FUNCTION_BLOCK "640_Rollenbahnen"   // FB640, SCL
{ S7_Optimized_Access := 'FALSE' }
AUTHOR : DJonas
VERSION : 0.1
   VAR_INPUT
      Notaus : Bool;
      Betriebsbereit : Bool;
      Start : Bool;
      StartRB : Bool;
      "630_Grundstellung" : Bool;
      i_s_grün : Bool;
      i_s_blau : Bool;
      i_Farbe_Code : Int;
   END_VAR
   VAR_OUTPUT
      o_RB_Frei : Bool;
      o_kontrolliert : Bool;
   END_VAR
   VAR_IN_OUT
      o_Farbsensor_Code : Int;
      o_kontrolle_fehler : Bool;
   END_VAR
   VAR
      RB9001_belegt : Bool;
      RB9002_belegt : Bool;
      RB9003_Belegt : Bool;
      Fehler : Bool;
      Neustart : TP;
      RB9001 : "641_Rollenbahn";
      RB9002 : "641_Rollenbahn";
      RB9003 : "641_Rollenbahn";
      B9002_RB9001_ntrig : "1001_300-ntrig-scl";
      B9004_RB9002_ntrig : "1001_300-ntrig-scl";
      B9006_RB9003_ntrig : "1001_300-ntrig-scl";
   END_VAR
BEGIN
   // Neustart Rollenbahn 2s laufen lassen um evtl. vorhandene Paletten vor einen Sensor zu fördern
   #Neustart(IN := #Notaus AND #Betriebsbereit, PT := T#2s);

   // Fehler Überbabe ohne Palette
   IF #StartRB AND NOT ("B9001_RB9001" OR "B9002_RB9001") THEN
       #Fehler := 1;
   ELSIF "B9006_RB9003" THEN
       #Fehler := 0;
   END_IF; 

   // Farbcode der Sensoren erstellen
   IF #i_s_blau THEN
       #o_Farbsensor_Code := 1;
   ELSIF #i_s_grün THEN
       #o_Farbsensor_Code := 2;
   ELSE
       #o_Farbsensor_Code := 0;
   END_IF;

   // Erkennung falsche Farbe auf Palette
   // ((#i_s_blau OR #i_s_grün) AND NOT (#i_Farbe_Code = #o_Farbsensor_Code))
   IF #Fehler AND #Betriebsbereit THEN
       #o_kontrolle_fehler := 1;
   END_IF;
   (*
   IF #o_kontrolle_fehler AND #Start THEN
       #o_Farbsensor_Code := #i_Farbe_Code;
       #o_kontrolliert := 1;
       #o_kontrolle_fehler := 0;
       #o_RB_Frei := 0;
       #Fehler := 0;
       RETURN;
   END_IF; *)

   // Kontrolle OK
   #o_kontrolliert := ((#i_s_blau OR #i_s_grün) AND (#i_Farbe_Code = #o_Farbsensor_Code)) OR #RB9003_Belegt OR #Fehler;

   // trigger für Stop Rollenbahn
   #B9002_RB9001_ntrig(IN := "B9002_RB9001" OR #Neustart.Q);
   #B9004_RB9002_ntrig(IN := "B9004_RB9002" OR #Neustart.Q);
   #B9006_RB9003_ntrig(IN := "B9006_RB9003" OR #Neustart.Q);

   // Ausgabe Rollenbahn 9001 und 9002 frei
   #o_RB_Frei := NOT #RB9001.belegt OR NOT #RB9002.belegt OR NOT #RB9003.belegt ;

   // Ansteuerung Rollenbahnen
   #RB9001(i_Start1:=(#StartRB OR #Neustart.Q),
           i_Start2:=("B9001_RB9001" OR "B9002_RB9001") AND #"630_Grundstellung",
           i_Stop:=#B9002_RB9001_ntrig.OUT OR (NOT #Betriebsbereit AND #"630_Grundstellung"),
           i_Halt:= NOT #"630_Grundstellung",
           i_NotHalt:=#Notaus,
           Output=>"RB9001",
           belegt:=#RB9001_belegt);

   #RB9002(i_Start1 := #Neustart.Q,
           i_Start2 := (("B9002_RB9001" AND #RB9001.Output) OR "B9003_RB9002"),
           i_Stop := #B9004_RB9002_ntrig.OUT OR (NOT #Betriebsbereit AND #"630_Grundstellung" AND #o_RB_Frei),
           i_NotHalt := #Notaus,
           Output => "RB9002",
           belegt := #RB9002_belegt);

   #RB9003(i_Start1:=#Neustart.Q,
           i_Start2:=("B9004_RB9002" OR "B9005_RB9003"),
           i_Stop:=#B9006_RB9003_ntrig.OUT OR (NOT #Betriebsbereit AND #"630_Grundstellung" AND #o_RB_Frei),
           i_NotHalt:=#Notaus,
           Output=>"RB9003",
           belegt:=#RB9003_Belegt);
END_FUNCTION_BLOCK

FUNCTION_BLOCK "641_Rollenbahn"   // FB641, SCL
{ S7_Optimized_Access := 'FALSE' }
VERSION : 0.1
   VAR_INPUT
      i_Start1 : Bool;
      i_Start2 : Bool;
      i_Halt : Bool;
      i_Stop : Bool;
      i_NotHalt : Bool;
   END_VAR
   VAR_OUTPUT
      Output : Bool;
   END_VAR
   VAR_IN_OUT
      belegt : Bool;
   END_VAR
BEGIN

   // Rollenbahn belegt setzen
   IF #i_Start1 OR #i_Start2 THEN
       #belegt := 1;
   END_IF;

   // Rollenbahn belegt entfernen
   IF #i_Stop OR NOT #i_NotHalt THEN
       #belegt := 0;
   END_IF;

   // Ausgang setzen wenn Rollenbahn belegt, kein Halt und kein Nothalt(zusätzlicher Schutz)
   #Output := #belegt AND #i_NotHalt AND  NOT #i_Halt;
END_FUNCTION_BLOCK

FUNCTION_BLOCK "1001_300-ntrig-scl"   // FB1001, SCL
{ S7_Optimized_Access := 'FALSE' }
VERSION : 0.1
   VAR_INPUT
      IN : Bool;
   END_VAR
   VAR_OUTPUT
      OUT : Bool;
   END_VAR
   VAR
      Merker : Bool;
   END_VAR
BEGIN
   #OUT := #Merker AND NOT #IN;
   #Merker := #IN;
END_FUNCTION_BLOCK

// ===== library: MasterCopy "RB_TB_einfach" =====

FUNCTION_BLOCK "RB_TB_einfach"   // FB101, GRAPH
{ S7_Optimized_Access := 'FALSE' }
VERSION : 0.1
// Einfacher Steuerbaustein RB / TB 
// Sensor Anfang / Ende  NO
   VAR_INPUT
      INIT_SQ : Bool := false;   // Kette in Initialzustand versetzen
      A_EIN : Bool;
      A_NOT_HALT : Bool;
      Nachfolgendes_Agg_frei : Bool;
      Sensor_vorheriges_Agg : Bool;
      Sensor_Anfang : Bool;   // Öffner
      Sensor_Ende : Bool;   // Öffner
   END_VAR
   VAR_OUTPUT
      Schritt_Nummer : Int;
      Aggregat : Bool;
      Aggregat_frei : Bool;
   END_VAR
   VAR
      HM_FLAM : Array[1..8] of Bool;
      Flanke : Array[1..8] of Bool;
      HM_Agg_Frei : Bool;
      HM_belegt : Bool;
      SWITCH : Array[0..0] of DWord;
      SW_SQTS : Array[0..6] of Byte;
      SW_ADDR : Word := 16#C;
      G7T_0 : GraphTransition;
      G7S_0 : GraphStep;
      PRE_CRIT : Array[0..1] of DWord;
      POST_CRIT : Array[0..0] of DWord;
      TVX : Array[0..2] of Byte;
      TTX : Array[0..2] of Byte;
      TSX : Array[0..2] of Byte;
      S00X : Array[0..2] of Byte;
      SOFFX : Array[0..2] of Byte;
      SONX : Array[0..2] of Byte;
      SAX : Array[0..2] of Byte;
      SERRX : Array[0..7] of Byte;
      SMX : Array[0..7] of Byte;
      S0X : Array[0..7] of Byte;
      S1X : Array[0..7] of Byte;
      S_DISPLAY : Int;   // Interne Anzeige des Ausgangsparameters S_NO
      S_SEL_OLD : Int;   // Vorheriger Wert an S_SEL
      S_DISPIDX : Byte;   // Index des Schritts, der an S_NO anliegt
      T_DISPIDX : Byte;   // Index der Transition, die an T_NO anliegt
      MOPEDGE : Struct
         AUTO : Bool := false;
         MAN : Bool := false;
         TAP : Bool := false;
         TOP : Bool := false;
         ACK_S : Bool := false;
         REG_S : Bool := false;
         T_PREV : Bool := false;
         T_NEXT : Bool := false;
         LOCK : Bool := false;
         SUP : Bool := false;
         ACKREQ : Bool := false;
         SSKIP : Bool := false;
         OFF : Bool := false;
         INIT : Bool := false;
         HALT : Bool := false;
         TMS_HALT : Bool := false;
         OPS_ZERO : Bool := false;
         SACT_DISP : Bool := false;
         SEF_DISP : Bool := false;
         SALL_DISP : Bool := false;
         S_PREV : Bool := false;
         S_NEXT : Bool := false;
         S_SELOK : Bool := false;
         S_ON : Bool := false;
         S_OFF : Bool := false;
         T_PUSH : Bool := false;
         REG : Bool := false;
         ACK : Bool := false;
         IL_PERM : Bool := false;
         T_PERM : Bool := false;
         ILP_MAN : Bool := false;
      END_STRUCT;
      MOP : Struct   // Betriebsart
         AUTO : Bool := true;   // Zustand: Automatischer Betrieb
         MAN : Bool := false;   // Zustand: Handbetrieb
         TAP : Bool := false;   // Zustand: Halbautomatisch/Weiterschalten mit Transition
         TOP : Bool := false;   // Zustand: Halbautomatisch/Ignoriere Transition
         ACK_S : Bool := false;   // Anforderung: Schritt quittieren, der an Parameter S_NO anliegt
         REG_S : Bool := false;   // Anforderung: Schritt registrieren, der an Parameter S_NO anliegt
         T_PREV : Bool := false;   // Anforderung: Vorherige gültige Transition am Parameter T_NO ausgeben
         T_NEXT : Bool := false;   // Anforderung: Nächste gültige Transition am Parameter T_NO ausgeben
         LOCK : Bool := true;   // Zustand: Interlockbearbeitung aktiviert
         SUP : Bool := true;   // Zustand: Supervisionsbearbeitung aktiviert
         ACKREQ : Bool := false;   // Zustand: Quittierung erforderlich
         SSKIP : Bool := false;   // Zustand: "Schritte überspringen" aktiviert
         OFF : Bool := false;   // Anforderung: Alle Schritte deaktivieren
         INIT : Bool := true;   // Anforderung: Kette in Initialzustand schalten
         HALT : Bool := false;   // Zustand: Kette schaltet nicht weiter
         TMS_HALT : Bool := false;   // Zustand: Alle internen Zeiten angehalten
         OPS_ZERO : Bool := false;   // Zustand: Alle mit N, L, D bearbeitete Operanden auf 0 gesetzt
         SACT_DISP : Bool := true;   // Zustand: Nur aktive Schritte anzeigen
         SEF_DISP : Bool := false;   // Zustand: Nur fehlerhafte und gestörte Schritte anzeigen
         SALL_DISP : Bool := false;   // Zustand: Alle Schritte anzeigen
         S_PREV : Bool := false;   // Anforderung: Vorherigen Schritt am Parameter S_NO ausgeben
         S_NEXT : Bool := false;   // Anforderung: Nächsten Schritt am Parameter S_NO ausgeben
         S_SELOK : Bool := false;   // Anforderung: Schrittnummer, die am Parameter S_SEL anliegt, am Parameter S_NO ausgeben
         S_ON : Bool := false;   // Anforderung: Schritt aktivieren, der am Parameter S_NO anliegt
         S_OFF : Bool := false;   // Anforderung: Schritt deaktivieren, der am Parameter S_NO anliegt
         T_PUSH : Bool := false;   // Anforderung: Schaltfreigabe für Transition
         REG : Bool := false;   // Anforderung: Alle Interlock- und Supervisionsfehler registrieren
         ACK : Bool := false;   // Anforderung: Alle Interlock- und Supervisionsfehler quittieren
         IL_PERM : Bool := false;   // Zustand: Permanente Bearbeitung aller Interlocks
         T_PERM : Bool := false;   // Zustand: Permanente Bearbeitung aller Transitionen
         ILP_MAN : Bool := false;   // Zustand: Permanente Bearbeitung aller Interlocks im Handbetrieb
      END_STRUCT;
      TICKS : Struct   // Zeittakte
         DELTA : Time := T#0ms;   // Zeitdifferenz zwischen zwei Zyklen
         OLD : Time := T#0ms;   // 10 ms Taktzählerstand im letzten Zyklus
         NEW : Time := T#0ms;   // 10 ms Taktzählerstand in diesem Zyklus
      END_STRUCT;
      SQ_FLAGS : Struct   // Kettenmerker
         ERR_FLT : Bool := false;   // Sammelfehler Interlock und Supervision
         ERROR : Bool := false;   // Sammelfehler Interlock
         FAULT : Bool := false;   // Sammelfehler Supervision
         RT_FAIL : Bool := false;   // Laufzeitfehler
         NO_SNO : Bool := false;   // Angeforderte Schrittnummer nicht gefunden
         NF_OFL : Bool := false;   // Überlauf: Zu viele Anforderungen ON oder OFF
         SA_OFL : Bool := false;   // Überlauf: Zu viele Schritte aktiv
         TV_OFL : Bool := false;   // Überlauf: Zu viele gültige Transitionen
         MSG_OFL : Bool := false;   // Überlauf: Nicht genügend Systemressourcen fü ALARM_S
         NO_SWI : Bool := false;   // Nicht Schalten in diesem Zyklus
         CYC_OP : Bool := false;   // Zyklische Bearbeitung der Kette nach Initialisierung
         AS_MSG : Bool := true;   // Meldungen zur Laufzeit durch Anweisung aktiviert oder deaktiviert
         AS_SEND : Bool := false;   // Meldungen von WR_USMSG senden oder nur in Diagnosepuffer eintragen
         SQ_BUSY : Bool := false;   // Interner Flankenmerker für Vorgangsbearbeitung
         SA_BUSY : Bool := false;   // Interner Flankenmerker für Vorgangsbearbeitung
         AS_SIG : Bool := false;   // Flankenmerker für Meldungen von Alarm_S und Alarm_SQ
      END_STRUCT;
      S_PTR : DWord := 16#450;
      S_PTR2 : DWord := 16#0;
      S_PTR3 : DWord := 16#D50;
      S_PTR4 : DWord := 16#D10;
      T_PTR : DWord := 16#CD0;
      C_AR2 : DWord := 16#0;
      M_FBDB : DWord := 16#640000;
      M_SNO : Word := 16#4;
      M_EVID : Word := 16#0;
      M_EVIL : C_Alarm_s;
      M_EVSV : C_Alarm_s;
      M_EV : DWord := 16#C30;
      CRIT : Array[0..31] of Bool;
      S_START : Byte := 16#0;
      S_IDX : Byte := 16#0;
      S_INT : Int := 72;
      S_TMP : Byte := 16#0;
      T_START : Byte := 16#0;
      T_IDX : Byte := 16#0;
      T_TMP : Byte := 16#0;
      T_TMP2 : Byte := 16#00;
      TV_POT : Byte := 16#02;
      RETURN1 : Byte := 16#0;
      RETURN2 : Byte := 16#0;
      SINI : Array[0..2] of Byte;
      LSTT : Array[0..6] of Byte;
      ATAJ : Array[0..6] of Byte;
      ATAB : Array[0..6] of Byte;
      PSTT : Array[0..6] of Byte;
      NSTT : Array[0..6] of Byte;
      ASSJ : Array[0..6] of Byte;
      ASSB : Array[0..6] of Byte;
      PTTS : Array[0..6] of Byte;
      NTTS : Array[0..6] of Byte;
      PRE_CNT : Word := 16#2;
      POST_CNT : Word := 16#1;
      ADR_COND : Word := 16#0;
      MAX_TVAL : Byte := 16#1;
      MAX_SACT : Byte := 16#1;
      MAX_CRIT : Byte := 16#4;
      T_CNT : Byte := 16#6;
      SUP_CNT : Byte := 16#0;
      LOCK_CNT : Byte := 16#5;
      S_CNT : Byte := 16#6;
      SQ_CNT : Byte := 16#1;
      PRS_INPAR : DWord := 16#40000000;
      PRS_OUTPAR : DWord := 16#0;
      GC_FLAGS : Struct
         T_MACH : Byte := 16#EB;
         COND_ED : Byte := 16#E2;
         W_LEVEL : Byte := 16#D5;
         FB_IF : Byte := 16#FA;
         AS_MSG : Word := 16#404;
         SSB : Word := 16#108;
         DILG : Word := 16#27E;
         ADDR_T0 : Word := 16#1A;
         CRIT_AVAIL : Bool := false;
         SSKIP_AVAIL : Bool := true;
         SSKIP_ON : Bool := false;
         ACK_REQ : Bool := false;
         SYNC_AVAIL : Bool := true;
         ILP_MAN : Bool := false;
         SWM_LOCKED : Bool := false;
         SAVE_SW : Bool := true;
      END_STRUCT;
      G7_FBMARK : Byte := 16#3C;
      G7_RELEASE : Byte := 16#3C;
      G7_ID2 : Byte := 16#37;
      G7_ID1 : Byte := 16#47;
   END_VAR
   // SW_SQTS[0] := 16#1;
   // TVX[0] := 16#1;
   // TTX[0] := 16#1;
   // TSX[0] := 16#1;
   // S00X[0] := 16#1;
   // SOFFX[0] := 16#1;
   // SONX[0] := 16#1;
   // SAX[0] := 16#1;
   // SERRX[0] := 16#1;
   // SMX[0] := 16#1;
   // S0X[0] := 16#1;
   // S1X[0] := 16#1;
   // SINI[0] := 16#2;
   // SINI[1] := 16#1;
   // SINI[2] := 0;
   // LSTT[0] := 0;
   // LSTT[1] := 0;
   // LSTT[2] := 0;
   // LSTT[3] := 0;
   // LSTT[4] := 0;
   // LSTT[5] := 0;
   // ATAJ[0] := 0;
   // ATAJ[1] := 16#1;
   // ATAJ[2] := 16#2;
   // ATAJ[3] := 16#3;
   // ATAJ[4] := 16#4;
   // ATAJ[5] := 16#5;
   // ATAB[0] := 0;
   // ATAB[1] := 16#1;
   // ATAB[2] := 16#2;
   // ATAB[3] := 16#3;
   // ATAB[4] := 16#4;
   // ATAB[5] := 16#5;
   // PSTT[0] := 0;
   // PSTT[1] := 16#1;
   // PSTT[2] := 16#2;
   // PSTT[3] := 16#3;
   // PSTT[4] := 16#4;
   // PSTT[5] := 16#5;
   // NSTT[0] := 16#1;
   // NSTT[1] := 16#2;
   // NSTT[2] := 16#3;
   // NSTT[3] := 16#4;
   // NSTT[4] := 16#5;
   // NSTT[5] := 16#6;
   // ASSJ[0] := 0;
   // ASSJ[1] := 16#1;
   // ASSJ[2] := 16#2;
   // ASSJ[3] := 16#3;
   // ASSJ[4] := 16#4;
   // ASSJ[5] := 16#5;
   // ASSB[0] := 0;
   // ASSB[1] := 16#1;
   // ASSB[2] := 16#2;
   // ASSB[3] := 16#3;
   // ASSB[4] := 16#4;
   // ASSB[5] := 16#5;
   // PTTS[0] := 0;
   // PTTS[2] := 16#1;
   // PTTS[3] := 16#2;
   // PTTS[4] := 16#3;
   // PTTS[5] := 16#4;
   // NTTS[0] := 0;
   // NTTS[1] := 16#1;
   // NTTS[2] := 16#2;
   // NTTS[3] := 16#3;
   // NTTS[4] := 16#4;
   // NTTS[5] := 16#5;
   // LSTT[6] := 16#1;
   // ATAJ[6] := 16#6;
   // ATAB[6] := 16#6;
   // PSTT[6] := 16#6;
   // NSTT[6] := 16#1;
   // ASSJ[6] := 16#6;
   // ASSB[6] := 16#6;
   // PTTS[6] := 16#5;
   // NTTS[6] := 16#6;
BEGIN
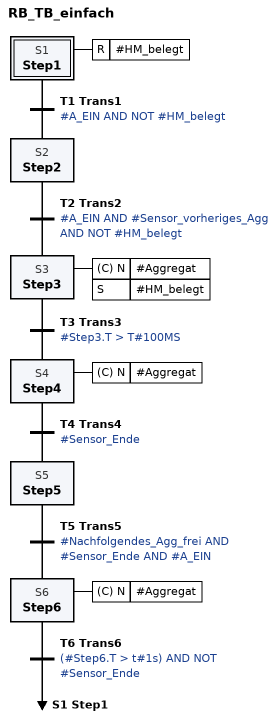
   // permanent pre-instructions
   NETWORK 1
      #HM_Agg_Frei := NOT #HM_belegt;
      #Aggregat_frei := NOT #HM_belegt;
   NETWORK 2
   TITLE = Ausgabe Schrittnummer
      #Schritt_Nummer := #S_DISPLAY;

   // sequencer 1
   INITIAL_STEP Step1:   // S1
      interlock C := NOT #A_NOT_HALT;
      // Warten auf Start
              R    #HM_belegt
   END_STEP
   TRANSITION Trans1 FROM Step1 TO Step2   // T1
      := #A_EIN AND NOT #HM_belegt;
   END_TRANSITION
   STEP Step4:   // S4
      interlock C := NOT #A_NOT_HALT;
      // Einfahrt bis Ende
      (C)     N    #Aggregat
   END_STEP
   TRANSITION Trans4 FROM Step4 TO Step5   // T4
      := #Sensor_Ende;
   END_TRANSITION
   STEP Step5:   // S5
      interlock C := NOT #A_NOT_HALT;
      // Warten auf Ausfahrt
   END_STEP
   TRANSITION Trans5 FROM Step5 TO Step6   // T5
      := #Nachfolgendes_Agg_frei AND #Sensor_Ende AND #A_EIN;
   END_TRANSITION
   STEP Step6:   // S6
      interlock C := NOT #A_NOT_HALT;
      // Ausfahrt bis Ende
      (C)     N    #Aggregat
   END_STEP
   TRANSITION Trans6 FROM Step6 TO Step1   // T6, jump
      := (#Step6.T > t#1s) AND NOT #Sensor_Ende;
   END_TRANSITION
   STEP Step3:   // S3
      interlock C := NOT #A_NOT_HALT;
      // Einfahrt Start
      (C)     N    #Aggregat
              S    #HM_belegt
   END_STEP
   TRANSITION Trans3 FROM Step3 TO Step4   // T3
      := #Step3.T > T#100MS;
   END_TRANSITION
   STEP Step2:   // S2
   END_STEP
   TRANSITION Trans2 FROM Step2 TO Step3   // T2
      := #A_EIN AND #Sensor_vorheriges_Agg AND NOT #HM_belegt;
   END_TRANSITION
END_FUNCTION_BLOCK

// ===== library: MasterCopy "Baustein_1" =====

FUNCTION_BLOCK "Baustein_1"   // FB2222, GRAPH
{ S7_Optimized_Access := 'FALSE' }
VERSION : 0.1
   VAR_INPUT
      INIT_SQ : Bool := false;   // Kette in Initialzustand versetzen
      A_EIN : Bool;
      A_NOT_HALT : Bool;
      Nachfolgendes_Agg_frei : Bool;
      Sensor_vorheriges_Agg : Bool;
      Sensor_Anfang : Bool;   // Öffner
      Sensor_Ende : Bool;   // Öffner
   END_VAR
   VAR_OUTPUT
      Schritt_Nummer : Int;
      Aggregat : Bool;
      Aggregat_frei : Bool;
   END_VAR
   VAR
      HM_FLAM : Array[1..8] of Bool;
      Flanke : Array[1..8] of Bool;
      HM_Agg_Frei : Bool;
      HM_belegt : Bool;
      SWITCH : Array[0..0] of DWord;
      SW_SQTS : Array[0..6] of Byte;
      SW_ADDR : Word := 16#C;
      G7T_0 : GraphTransition;
      G7S_0 : GraphStep;
      PRE_CRIT : Array[0..1] of DWord;
      POST_CRIT : Array[0..0] of DWord;
      TVX : Array[0..2] of Byte;
      TTX : Array[0..2] of Byte;
      TSX : Array[0..2] of Byte;
      S00X : Array[0..2] of Byte;
      SOFFX : Array[0..2] of Byte;
      SONX : Array[0..2] of Byte;
      SAX : Array[0..2] of Byte;
      SERRX : Array[0..7] of Byte;
      SMX : Array[0..7] of Byte;
      S0X : Array[0..7] of Byte;
      S1X : Array[0..7] of Byte;
      S_DISPLAY : Int;   // Interne Anzeige des Ausgangsparameters S_NO
      S_SEL_OLD : Int;   // Vorheriger Wert an S_SEL
      S_DISPIDX : Byte;   // Index des Schritts, der an S_NO anliegt
      T_DISPIDX : Byte;   // Index der Transition, die an T_NO anliegt
      MOPEDGE : Struct
         AUTO : Bool := false;
         MAN : Bool := false;
         TAP : Bool := false;
         TOP : Bool := false;
         ACK_S : Bool := false;
         REG_S : Bool := false;
         T_PREV : Bool := false;
         T_NEXT : Bool := false;
         LOCK : Bool := false;
         SUP : Bool := false;
         ACKREQ : Bool := false;
         SSKIP : Bool := false;
         OFF : Bool := false;
         INIT : Bool := false;
         HALT : Bool := false;
         TMS_HALT : Bool := false;
         OPS_ZERO : Bool := false;
         SACT_DISP : Bool := false;
         SEF_DISP : Bool := false;
         SALL_DISP : Bool := false;
         S_PREV : Bool := false;
         S_NEXT : Bool := false;
         S_SELOK : Bool := false;
         S_ON : Bool := false;
         S_OFF : Bool := false;
         T_PUSH : Bool := false;
         REG : Bool := false;
         ACK : Bool := false;
         IL_PERM : Bool := false;
         T_PERM : Bool := false;
         ILP_MAN : Bool := false;
      END_STRUCT;
      MOP : Struct   // Betriebsart
         AUTO : Bool := true;   // Zustand: Automatischer Betrieb
         MAN : Bool := false;   // Zustand: Handbetrieb
         TAP : Bool := false;   // Zustand: Halbautomatisch/Weiterschalten mit Transition
         TOP : Bool := false;   // Zustand: Halbautomatisch/Ignoriere Transition
         ACK_S : Bool := false;   // Anforderung: Schritt quittieren, der an Parameter S_NO anliegt
         REG_S : Bool := false;   // Anforderung: Schritt registrieren, der an Parameter S_NO anliegt
         T_PREV : Bool := false;   // Anforderung: Vorherige gültige Transition am Parameter T_NO ausgeben
         T_NEXT : Bool := false;   // Anforderung: Nächste gültige Transition am Parameter T_NO ausgeben
         LOCK : Bool := true;   // Zustand: Interlockbearbeitung aktiviert
         SUP : Bool := true;   // Zustand: Supervisionsbearbeitung aktiviert
         ACKREQ : Bool := false;   // Zustand: Quittierung erforderlich
         SSKIP : Bool := false;   // Zustand: "Schritte überspringen" aktiviert
         OFF : Bool := false;   // Anforderung: Alle Schritte deaktivieren
         INIT : Bool := true;   // Anforderung: Kette in Initialzustand schalten
         HALT : Bool := false;   // Zustand: Kette schaltet nicht weiter
         TMS_HALT : Bool := false;   // Zustand: Alle internen Zeiten angehalten
         OPS_ZERO : Bool := false;   // Zustand: Alle mit N, L, D bearbeitete Operanden auf 0 gesetzt
         SACT_DISP : Bool := true;   // Zustand: Nur aktive Schritte anzeigen
         SEF_DISP : Bool := false;   // Zustand: Nur fehlerhafte und gestörte Schritte anzeigen
         SALL_DISP : Bool := false;   // Zustand: Alle Schritte anzeigen
         S_PREV : Bool := false;   // Anforderung: Vorherigen Schritt am Parameter S_NO ausgeben
         S_NEXT : Bool := false;   // Anforderung: Nächsten Schritt am Parameter S_NO ausgeben
         S_SELOK : Bool := false;   // Anforderung: Schrittnummer, die am Parameter S_SEL anliegt, am Parameter S_NO ausgeben
         S_ON : Bool := false;   // Anforderung: Schritt aktivieren, der am Parameter S_NO anliegt
         S_OFF : Bool := false;   // Anforderung: Schritt deaktivieren, der am Parameter S_NO anliegt
         T_PUSH : Bool := false;   // Anforderung: Schaltfreigabe für Transition
         REG : Bool := false;   // Anforderung: Alle Interlock- und Supervisionsfehler registrieren
         ACK : Bool := false;   // Anforderung: Alle Interlock- und Supervisionsfehler quittieren
         IL_PERM : Bool := false;   // Zustand: Permanente Bearbeitung aller Interlocks
         T_PERM : Bool := false;   // Zustand: Permanente Bearbeitung aller Transitionen
         ILP_MAN : Bool := false;   // Zustand: Permanente Bearbeitung aller Interlocks im Handbetrieb
      END_STRUCT;
      TICKS : Struct   // Zeittakte
         DELTA : Time := T#0ms;   // Zeitdifferenz zwischen zwei Zyklen
         OLD : Time := T#0ms;   // 10 ms Taktzählerstand im letzten Zyklus
         NEW : Time := T#0ms;   // 10 ms Taktzählerstand in diesem Zyklus
      END_STRUCT;
      SQ_FLAGS : Struct   // Kettenmerker
         ERR_FLT : Bool := false;   // Sammelfehler Interlock und Supervision
         ERROR : Bool := false;   // Sammelfehler Interlock
         FAULT : Bool := false;   // Sammelfehler Supervision
         RT_FAIL : Bool := false;   // Laufzeitfehler
         NO_SNO : Bool := false;   // Angeforderte Schrittnummer nicht gefunden
         NF_OFL : Bool := false;   // Überlauf: Zu viele Anforderungen ON oder OFF
         SA_OFL : Bool := false;   // Überlauf: Zu viele Schritte aktiv
         TV_OFL : Bool := false;   // Überlauf: Zu viele gültige Transitionen
         MSG_OFL : Bool := false;   // Überlauf: Nicht genügend Systemressourcen fü ALARM_S
         NO_SWI : Bool := false;   // Nicht Schalten in diesem Zyklus
         CYC_OP : Bool := false;   // Zyklische Bearbeitung der Kette nach Initialisierung
         AS_MSG : Bool := true;   // Meldungen zur Laufzeit durch Anweisung aktiviert oder deaktiviert
         AS_SEND : Bool := false;   // Meldungen von WR_USMSG senden oder nur in Diagnosepuffer eintragen
         SQ_BUSY : Bool := false;   // Interner Flankenmerker für Vorgangsbearbeitung
         SA_BUSY : Bool := false;   // Interner Flankenmerker für Vorgangsbearbeitung
         AS_SIG : Bool := false;   // Flankenmerker für Meldungen von Alarm_S und Alarm_SQ
      END_STRUCT;
      S_PTR : DWord := 16#450;
      S_PTR2 : DWord := 16#0;
      S_PTR3 : DWord := 16#D50;
      S_PTR4 : DWord := 16#D10;
      T_PTR : DWord := 16#CD0;
      C_AR2 : DWord := 16#0;
      M_FBDB : DWord := 16#8AE0000;
      M_SNO : Word := 16#4;
      M_EVID : Word := 16#0;
      M_EVIL : C_Alarm_s;
      M_EVSV : C_Alarm_s;
      M_EV : DWord := 16#C30;
      CRIT : Array[0..31] of Bool;
      S_START : Byte := 16#0;
      S_IDX : Byte := 16#0;
      S_INT : Int := 72;
      S_TMP : Byte := 16#0;
      T_START : Byte := 16#0;
      T_IDX : Byte := 16#0;
      T_TMP : Byte := 16#0;
      T_TMP2 : Byte := 16#00;
      TV_POT : Byte := 16#02;
      RETURN1 : Byte := 16#0;
      RETURN2 : Byte := 16#0;
      SINI : Array[0..2] of Byte;
      LSTT : Array[0..6] of Byte;
      ATAJ : Array[0..6] of Byte;
      ATAB : Array[0..6] of Byte;
      PSTT : Array[0..6] of Byte;
      NSTT : Array[0..6] of Byte;
      ASSJ : Array[0..6] of Byte;
      ASSB : Array[0..6] of Byte;
      PTTS : Array[0..6] of Byte;
      NTTS : Array[0..6] of Byte;
      PRE_CNT : Word := 16#2;
      POST_CNT : Word := 16#1;
      ADR_COND : Word := 16#0;
      MAX_TVAL : Byte := 16#1;
      MAX_SACT : Byte := 16#1;
      MAX_CRIT : Byte := 16#4;
      T_CNT : Byte := 16#6;
      SUP_CNT : Byte := 16#0;
      LOCK_CNT : Byte := 16#5;
      S_CNT : Byte := 16#6;
      SQ_CNT : Byte := 16#1;
      PRS_INPAR : DWord := 16#40000000;
      PRS_OUTPAR : DWord := 16#0;
      GC_FLAGS : Struct
         T_MACH : Byte := 16#EB;
         COND_ED : Byte := 16#E2;
         W_LEVEL : Byte := 16#D5;
         FB_IF : Byte := 16#FA;
         AS_MSG : Word := 16#404;
         SSB : Word := 16#108;
         DILG : Word := 16#27E;
         ADDR_T0 : Word := 16#1A;
         CRIT_AVAIL : Bool := false;
         SSKIP_AVAIL : Bool := true;
         SSKIP_ON : Bool := false;
         ACK_REQ : Bool := false;
         SYNC_AVAIL : Bool := true;
         ILP_MAN : Bool := false;
         SWM_LOCKED : Bool := false;
         SAVE_SW : Bool := true;
      END_STRUCT;
      G7_FBMARK : Byte := 16#3C;
      G7_RELEASE : Byte := 16#3C;
      G7_ID2 : Byte := 16#37;
      G7_ID1 : Byte := 16#47;
   END_VAR
   // SW_SQTS[0] := 16#1;
   // TVX[0] := 16#1;
   // TTX[0] := 16#1;
   // TSX[0] := 16#1;
   // S00X[0] := 16#1;
   // SOFFX[0] := 16#1;
   // SONX[0] := 16#1;
   // SAX[0] := 16#1;
   // SERRX[0] := 16#1;
   // SMX[0] := 16#1;
   // S0X[0] := 16#1;
   // S1X[0] := 16#1;
   // SINI[0] := 16#2;
   // SINI[1] := 16#1;
   // SINI[2] := 0;
   // LSTT[0] := 0;
   // LSTT[1] := 0;
   // LSTT[2] := 0;
   // LSTT[3] := 0;
   // LSTT[4] := 0;
   // LSTT[5] := 0;
   // LSTT[6] := 16#1;
   // ATAJ[0] := 0;
   // ATAJ[1] := 16#1;
   // ATAJ[2] := 16#2;
   // ATAJ[3] := 16#3;
   // ATAJ[4] := 16#4;
   // ATAJ[5] := 16#5;
   // ATAJ[6] := 16#6;
   // ATAB[0] := 0;
   // ATAB[1] := 16#1;
   // ATAB[2] := 16#2;
   // ATAB[3] := 16#3;
   // ATAB[4] := 16#4;
   // ATAB[5] := 16#5;
   // ATAB[6] := 16#6;
   // PSTT[0] := 0;
   // PSTT[1] := 16#1;
   // PSTT[2] := 16#2;
   // PSTT[3] := 16#3;
   // PSTT[4] := 16#4;
   // PSTT[5] := 16#5;
   // PSTT[6] := 16#6;
   // NSTT[0] := 16#1;
   // NSTT[1] := 16#2;
   // NSTT[2] := 16#3;
   // NSTT[3] := 16#4;
   // NSTT[4] := 16#5;
   // NSTT[5] := 16#6;
   // NSTT[6] := 16#1;
   // ASSJ[0] := 0;
   // ASSJ[1] := 16#1;
   // ASSJ[2] := 16#2;
   // ASSJ[3] := 16#3;
   // ASSJ[4] := 16#4;
   // ASSJ[5] := 16#5;
   // ASSJ[6] := 16#6;
   // ASSB[0] := 0;
   // ASSB[1] := 16#1;
   // ASSB[2] := 16#2;
   // ASSB[3] := 16#3;
   // ASSB[4] := 16#4;
   // ASSB[5] := 16#5;
   // ASSB[6] := 16#6;
   // PTTS[0] := 0;
   // PTTS[2] := 16#1;
   // PTTS[3] := 16#2;
   // PTTS[4] := 16#3;
   // PTTS[5] := 16#4;
   // PTTS[6] := 16#5;
   // NTTS[0] := 0;
   // NTTS[1] := 16#1;
   // NTTS[2] := 16#2;
   // NTTS[3] := 16#3;
   // NTTS[4] := 16#4;
   // NTTS[5] := 16#5;
   // NTTS[6] := 16#6;
BEGIN
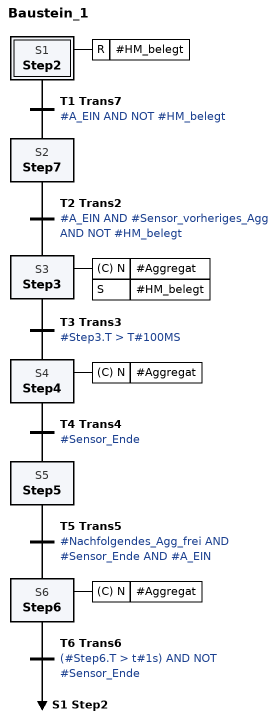
   // permanent pre-instructions
   NETWORK 1
      #HM_Agg_Frei := NOT #HM_belegt;
      #Aggregat_frei := NOT #HM_belegt;
   NETWORK 2
   TITLE = Ausgabe Schrittnummer
      #Schritt_Nummer := #S_DISPLAY;

   // sequencer 1
   INITIAL_STEP Step2:   // S1
      interlock C := NOT #A_NOT_HALT;
      // Warten auf Start
              R    #HM_belegt
   END_STEP
   TRANSITION Trans7 FROM Step2 TO Step7   // T1
      := #A_EIN AND NOT #HM_belegt;
   END_TRANSITION
   STEP Step4:   // S4
      interlock C := NOT #A_NOT_HALT;
      // Einfahrt bis Ende
      (C)     N    #Aggregat
   END_STEP
   TRANSITION Trans4 FROM Step4 TO Step5   // T4
      := #Sensor_Ende;
   END_TRANSITION
   STEP Step5:   // S5
      interlock C := NOT #A_NOT_HALT;
      // Warten auf Ausfahrt
   END_STEP
   TRANSITION Trans5 FROM Step5 TO Step6   // T5
      := #Nachfolgendes_Agg_frei AND #Sensor_Ende AND #A_EIN;
   END_TRANSITION
   STEP Step6:   // S6
      interlock C := NOT #A_NOT_HALT;
      // Ausfahrt bis Ende
      (C)     N    #Aggregat
   END_STEP
   TRANSITION Trans6 FROM Step6 TO Step2   // T6, jump
      := (#Step6.T > t#1s) AND NOT #Sensor_Ende;
   END_TRANSITION
   STEP Step3:   // S3
      interlock C := NOT #A_NOT_HALT;
      // Einfahrt Start
      (C)     N    #Aggregat
              S    #HM_belegt
   END_STEP
   TRANSITION Trans3 FROM Step3 TO Step4   // T3
      := #Step3.T > T#100MS;
   END_TRANSITION
   STEP Step7:   // S2
   END_STEP
   TRANSITION Trans2 FROM Step7 TO Step3   // T2
      := #A_EIN AND #Sensor_vorheriges_Agg AND NOT #HM_belegt;
   END_TRANSITION
END_FUNCTION_BLOCK

(* ===== HMI "HMI_RT_1" =====
system functions are stored by id; their names below are inferred from use
connection "HMI_Verbindung_1": MPI/DP, SIMATIC S7 300/400 MPI

HMI tags "Standard-Variablentabelle"
   "HochregallagerDB_Motors_Ein" : Bool = PLC HochregallagerDB.Motors_Ein AT %DB1.DBX10.1, 100 ms
   "HochregallagerDB_Automatik" : Bool = PLC HochregallagerDB.Automatik AT %DB1.DBX10.0, 100 ms
   "HochregallagerDB_Neue_Palette" : Bool = PLC HochregallagerDB.Neue_Palette AT %DB1.DBX10.2, 100 ms
   "Paketempfang_Rollenbahn_DB_Palette_auf_RB1" : Bool = PLC FB_Paketempfang_Rollenbahn_DB.Palette_auf_RB1 AT %DB2.DBX12.1, 100 ms
   "Paketempfang_Rollenbahn_DB_Palette_auf_RB2" : Bool = PLC FB_Paketempfang_Rollenbahn_DB.Palette_auf_RB2 AT %DB2.DBX12.2, 100 ms
   "Paketempfang_Rollenbahn_DB_Palette_auf_RB3" : Bool = PLC FB_Paketempfang_Rollenbahn_DB.Palette_auf_RB3 AT %DB2.DBX12.3, 100 ms
   "Paketempfang_Rollenbahn_DB_Farbe_RB2" : Int = PLC FB_Paketempfang_Rollenbahn_DB.Farbe_RB2 AT %DB2.DBW14, 100 ms
   "Paketempfang_Rollenbahn_DB_Farbe_RB3" : Int = PLC FB_Paketempfang_Rollenbahn_DB.Farbe_RB3 AT %DB2.DBW4, 100 ms
   "HochregallagerDB_Farbe" : Int = PLC HochregallagerDB.Farbe AT %DB1.DBW6, 100 ms
   "HochregallagerDB_HMI_X_Bewegung" : Int = PLC HochregallagerDB.HMI_X_Bewegung AT %DB1.DBW12, 100 ms
   "HochregallagerDB_HMI_Z_Bewegung" : Int = PLC HochregallagerDB.HMI_Z_Bewegung AT %DB1.DBW14, 100 ms
   "HochregallagerDB_Stappler_Aktuele_Farbe" : Int = PLC HochregallagerDB.Stappler_Aktuele_Farbe AT %DB1.DBW8, 100 ms
   "HochregallagerDB_Lagerplaetze{1}_Materialfarbe" : String[10] = PLC HochregallagerDB.Lagerplaetze[1].Materialfarbe AT %DB1.DBX26.0, 100 ms
   "HochregallagerDB_Lagerplaetze{1}_Materialfarbe_Nummer" : Int = PLC HochregallagerDB.Lagerplaetze[1].Materialfarbe_Nummer AT %DB1.DBW38, 100 ms
   "HochregallagerDB_Lagerplaetze{2}_Materialfarbe_Nummer" : Int = PLC HochregallagerDB.Lagerplaetze[2].Materialfarbe_Nummer AT %DB1.DBW62, 100 ms
   "HochregallagerDB_Lagerplaetze{3}_Materialfarbe_Nummer" : Int = PLC HochregallagerDB.Lagerplaetze[3].Materialfarbe_Nummer AT %DB1.DBW86, 100 ms
   "HochregallagerDB_Lagerplaetze{4}_Materialfarbe_Nummer" : Int = PLC HochregallagerDB.Lagerplaetze[4].Materialfarbe_Nummer AT %DB1.DBW110, 100 ms
   "HochregallagerDB_Lagerplaetze{5}_Materialfarbe_Nummer" : Int = PLC HochregallagerDB.Lagerplaetze[5].Materialfarbe_Nummer AT %DB1.DBW134, 100 ms
   "HochregallagerDB_Lagerplaetze{6}_Materialfarbe_Nummer" : Int = PLC HochregallagerDB.Lagerplaetze[6].Materialfarbe_Nummer AT %DB1.DBW158, 100 ms
   "HochregallagerDB_Lagerplaetze{7}_Materialfarbe_Nummer" : Int = PLC HochregallagerDB.Lagerplaetze[7].Materialfarbe_Nummer AT %DB1.DBW182, 100 ms
   "HochregallagerDB_Lagerplaetze{8}_Materialfarbe_Nummer" : Int = PLC HochregallagerDB.Lagerplaetze[8].Materialfarbe_Nummer AT %DB1.DBW206, 100 ms
   "HochregallagerDB_Lagerplaetze{9}_Materialfarbe_Nummer" : Int = PLC HochregallagerDB.Lagerplaetze[9].Materialfarbe_Nummer AT %DB1.DBW230, 100 ms
   "HochregallagerDB_Lagerplaetze{10}_Materialfarbe_Nummer" : Int = PLC HochregallagerDB.Lagerplaetze[10].Materialfarbe_Nummer AT %DB1.DBW254, 100 ms
   "HochregallagerDB_Lagerplaetze{11}_Materialfarbe_Nummer" : Int = PLC HochregallagerDB.Lagerplaetze[11].Materialfarbe_Nummer AT %DB1.DBW278, 100 ms
   "HochregallagerDB_Lagerplaetze{12}_Materialfarbe_Nummer" : Int = PLC HochregallagerDB.Lagerplaetze[12].Materialfarbe_Nummer AT %DB1.DBW302, 100 ms
   "HochregallagerDB_Lagerplaetze{13}_Materialfarbe_Nummer" : Int = PLC HochregallagerDB.Lagerplaetze[13].Materialfarbe_Nummer AT %DB1.DBW326, 100 ms
   "HochregallagerDB_Lagerplaetze{14}_Materialfarbe_Nummer" : Int = PLC HochregallagerDB.Lagerplaetze[14].Materialfarbe_Nummer AT %DB1.DBW350, 100 ms
   "HochregallagerDB_Lagerplaetze{15}_Materialfarbe_Nummer" : Int = PLC HochregallagerDB.Lagerplaetze[15].Materialfarbe_Nummer AT %DB1.DBW374, 100 ms
   "HochregallagerDB_Lagerplaetze{16}_Materialfarbe_Nummer" : Int = PLC HochregallagerDB.Lagerplaetze[16].Materialfarbe_Nummer AT %DB1.DBW398, 100 ms
   "HochregallagerDB_Lagerplaetze{17}_Materialfarbe_Nummer" : Int = PLC HochregallagerDB.Lagerplaetze[17].Materialfarbe_Nummer AT %DB1.DBW422, 100 ms
   "HochregallagerDB_Lagerplaetze{18}_Materialfarbe_Nummer" : Int = PLC HochregallagerDB.Lagerplaetze[18].Materialfarbe_Nummer AT %DB1.DBW446, 100 ms
   "HochregallagerDB_Lagerplaetze{19}_Materialfarbe_Nummer" : Int = PLC HochregallagerDB.Lagerplaetze[19].Materialfarbe_Nummer AT %DB1.DBW470, 100 ms
   "HochregallagerDB_Lagerplaetze{20}_Materialfarbe_Nummer" : Int = PLC HochregallagerDB.Lagerplaetze[20].Materialfarbe_Nummer AT %DB1.DBW494, 100 ms
   "HochregallagerDB_Lagerplaetze{21}_Materialfarbe_Nummer" : Int = PLC HochregallagerDB.Lagerplaetze[21].Materialfarbe_Nummer AT %DB1.DBW518, 100 ms
   "HochregallagerDB_Lagerplaetze{22}_Materialfarbe_Nummer" : Int = PLC HochregallagerDB.Lagerplaetze[22].Materialfarbe_Nummer AT %DB1.DBW542, 100 ms
   "HochregallagerDB_Lagerplaetze{23}_Materialfarbe_Nummer" : Int = PLC HochregallagerDB.Lagerplaetze[23].Materialfarbe_Nummer AT %DB1.DBW566, 100 ms
   "HochregallagerDB_Lagerplaetze{24}_Materialfarbe_Nummer" : Int = PLC HochregallagerDB.Lagerplaetze[24].Materialfarbe_Nummer AT %DB1.DBW590, 100 ms
   "HochregallagerDB_Lagerplaetze{25}_Materialfarbe_Nummer" : Int = PLC HochregallagerDB.Lagerplaetze[25].Materialfarbe_Nummer AT %DB1.DBW614, 100 ms
   "HochregallagerDB_Lagerplaetze{26}_Materialfarbe_Nummer" : Int = PLC HochregallagerDB.Lagerplaetze[26].Materialfarbe_Nummer AT %DB1.DBW638, 100 ms
   "HochregallagerDB_Lagerplaetze{27}_Materialfarbe_Nummer" : Int = PLC HochregallagerDB.Lagerplaetze[27].Materialfarbe_Nummer AT %DB1.DBW662, 100 ms
   "HochregallagerDB_Lagerplaetze{28}_Materialfarbe_Nummer" : Int = PLC HochregallagerDB.Lagerplaetze[28].Materialfarbe_Nummer AT %DB1.DBW686, 100 ms
   "HochregallagerDB_Lagerplaetze{29}_Materialfarbe_Nummer" : Int = PLC HochregallagerDB.Lagerplaetze[29].Materialfarbe_Nummer AT %DB1.DBW710, 100 ms
   "HochregallagerDB_Lagerplaetze{30}_Materialfarbe_Nummer" : Int = PLC HochregallagerDB.Lagerplaetze[30].Materialfarbe_Nummer AT %DB1.DBW734, 100 ms
   "HochregallagerDB_Lagerplaetze{31}_Materialfarbe_Nummer" : Int = PLC HochregallagerDB.Lagerplaetze[31].Materialfarbe_Nummer AT %DB1.DBW758, 100 ms
   "HochregallagerDB_Lagerplaetze{32}_Materialfarbe_Nummer" : Int = PLC HochregallagerDB.Lagerplaetze[32].Materialfarbe_Nummer AT %DB1.DBW782, 100 ms
   "HochregallagerDB_Lagerplaetze{33}_Materialfarbe_Nummer" : Int = PLC HochregallagerDB.Lagerplaetze[33].Materialfarbe_Nummer AT %DB1.DBW806, 100 ms
   "HochregallagerDB_Lagerplaetze{34}_Materialfarbe_Nummer" : Int = PLC HochregallagerDB.Lagerplaetze[34].Materialfarbe_Nummer AT %DB1.DBW830, 100 ms
   "HochregallagerDB_Lagerplaetze{35}_Materialfarbe_Nummer" : Int = PLC HochregallagerDB.Lagerplaetze[35].Materialfarbe_Nummer AT %DB1.DBW854, 100 ms
   "HochregallagerDB_Lagerplaetze{36}_Materialfarbe_Nummer" : Int = PLC HochregallagerDB.Lagerplaetze[36].Materialfarbe_Nummer AT %DB1.DBW878, 100 ms
   "HochregallagerDB_Lagerplaetze{37}_Materialfarbe_Nummer" : Int = PLC HochregallagerDB.Lagerplaetze[37].Materialfarbe_Nummer AT %DB1.DBW902, 100 ms
   "HochregallagerDB_Lagerplaetze{38}_Materialfarbe_Nummer" : Int = PLC HochregallagerDB.Lagerplaetze[38].Materialfarbe_Nummer AT %DB1.DBW926, 100 ms
   "HochregallagerDB_Lagerplaetze{39}_Materialfarbe_Nummer" : Int = PLC HochregallagerDB.Lagerplaetze[39].Materialfarbe_Nummer AT %DB1.DBW950, 100 ms
   "HochregallagerDB_Lagerplaetze{40}_Materialfarbe_Nummer" : Int = PLC HochregallagerDB.Lagerplaetze[40].Materialfarbe_Nummer AT %DB1.DBW974, 100 ms
   "HochregallagerDB_Lagerplaetze{41}_Materialfarbe_Nummer" : Int = PLC HochregallagerDB.Lagerplaetze[41].Materialfarbe_Nummer AT %DB1.DBW998, 100 ms
   "HochregallagerDB_Lagerplaetze{42}_Materialfarbe_Nummer" : Int = PLC HochregallagerDB.Lagerplaetze[42].Materialfarbe_Nummer AT %DB1.DBW1022, 100 ms
   "HochregallagerDB_Lagerplaetze{43}_Materialfarbe_Nummer" : Int = PLC HochregallagerDB.Lagerplaetze[43].Materialfarbe_Nummer AT %DB1.DBW1046, 100 ms
   "HochregallagerDB_Lagerplaetze{44}_Materialfarbe_Nummer" : Int = PLC HochregallagerDB.Lagerplaetze[44].Materialfarbe_Nummer AT %DB1.DBW1070, 100 ms
   "HochregallagerDB_Lagerplaetze{45}_Materialfarbe_Nummer" : Int = PLC HochregallagerDB.Lagerplaetze[45].Materialfarbe_Nummer AT %DB1.DBW1094, 100 ms
   "HochregallagerDB_Lagerplaetze{46}_Materialfarbe_Nummer" : Int = PLC HochregallagerDB.Lagerplaetze[46].Materialfarbe_Nummer AT %DB1.DBW1118, 100 ms
   "HochregallagerDB_Lagerplaetze{47}_Materialfarbe_Nummer" : Int = PLC HochregallagerDB.Lagerplaetze[47].Materialfarbe_Nummer AT %DB1.DBW1142, 100 ms
   "HochregallagerDB_Lagerplaetze{48}_Materialfarbe_Nummer" : Int = PLC HochregallagerDB.Lagerplaetze[48].Materialfarbe_Nummer AT %DB1.DBW1166, 100 ms
   "HochregallagerDB_Lagerplaetze{49}_Materialfarbe_Nummer" : Int = PLC HochregallagerDB.Lagerplaetze[49].Materialfarbe_Nummer AT %DB1.DBW1190, 100 ms
   "HochregallagerDB_Lagerplaetze{50}_Materialfarbe_Nummer" : Int = PLC HochregallagerDB.Lagerplaetze[50].Materialfarbe_Nummer AT %DB1.DBW1214, 100 ms
   "HochregallagerDB_Lagerplaetze{51}_Materialfarbe_Nummer" : Int = PLC HochregallagerDB.Lagerplaetze[51].Materialfarbe_Nummer AT %DB1.DBW1238, 100 ms
   "HochregallagerDB_Lagerplaetze{52}_Materialfarbe_Nummer" : Int = PLC HochregallagerDB.Lagerplaetze[52].Materialfarbe_Nummer AT %DB1.DBW1262, 100 ms
   "HochregallagerDB_Lagerplaetze{53}_Materialfarbe_Nummer" : Int = PLC HochregallagerDB.Lagerplaetze[53].Materialfarbe_Nummer AT %DB1.DBW1286, 100 ms
   "HochregallagerDB_Lagerplaetze{54}_Materialfarbe_Nummer" : Int = PLC HochregallagerDB.Lagerplaetze[54].Materialfarbe_Nummer AT %DB1.DBW1310, 100 ms
   "HochregallagerDB_Anzahl_Blau" : Int = PLC HochregallagerDB.Anzahl_Blau AT %DB1.DBW1314, 100 ms
   "HochregallagerDB_Anzahl_Gruen" : Int = PLC HochregallagerDB.Anzahl_Gruen AT %DB1.DBW1316, 100 ms
   "P10_START" : Bool = PLC P10_START AT %A0.3, 100 ms
   "P11_STOP" : Bool = PLC P11_STOP AT %A0.4, 100 ms
   "S2_START" : Bool = PLC S2_START AT %E0.2, 100 ms
   "HMI_Eingaben_DB_HMI_Start" : Bool = PLC HMI_Eingaben_DB.HMI_Start AT %DB8.DBX0.0, 100 ms
   "HMI_Eingaben_DB_HMI_Stop" : Bool = PLC HMI_Eingaben_DB.HMI_Stop AT %DB8.DBX0.1, 100 ms
   "HMI_Eingaben_DB_HMI_Not_Halt" : Bool = PLC HMI_Eingaben_DB.HMI_Not_Halt AT %DB8.DBX0.2, 100 ms
   "HMI_Eingaben_DB_HMI_Hauptschalter" : Bool = PLC HMI_Eingaben_DB.HMI_Hauptschalter AT %DB8.DBX0.3, 100 ms
   "P3_MS_GN" : Bool = PLC P3_MS_GN AT %A0.2, 100 ms
   "P2_MS_GE" : Bool = PLC P2_MS_GE AT %A0.1, 100 ms
   "P1_MS_RT" : Bool = PLC P1_MS_RT AT %A0.0, 100 ms
   "HMI_Eingaben_DB_HMI_Start_Anzeige" : Bool = PLC HMI_Eingaben_DB.HMI_Start_Anzeige AT %DB8.DBX0.4, 100 ms
   "HochregallagerDB_Lager_Voll" : Bool = PLC HochregallagerDB.Lager_Voll AT %DB1.DBX1322.5, 100 ms
   "HochregallagerDB_Warnung_Wenig_Freie_Plaetze" : Bool = PLC HochregallagerDB.Warnung_Wenig_Freie_Plaetze AT %DB1.DBX1322.4, 100 ms
   "HochregallagerDB_Stoerung_Aktiv" : Bool = PLC HochregallagerDB.Stoerung_Aktiv AT %DB1.DBX1322.2, 100 ms
   "P12_Anfahrwarnung" : Bool = PLC P12_Anfahrwarnung AT %A0.6, 100 ms
   "P8001_Warnung_Bewegung_1" : Bool = PLC P8001_Warnung_Bewegung_1 AT %A2.6, 100 ms
   "P8002_Warnung_Bewegung_2" : Bool = PLC P8002_Warnung_Bewegung_2 AT %A2.7, 100 ms
   "S2_START_1" : Bool AT %E0.3, 100 ms
   "HochregallagerDB_Anzahl_Unbekannte_Farbe" : Int = PLC HochregallagerDB.Anzahl_Unbekannte_Farbe AT %DB1.DBW1318, 100 ms

screen "Lafger" 1024x768
   Rectangle "Rechteck_57" at 596,12 size 47x36
      Appearance <- "HochregallagerDB_Lagerplaetze{53}_Materialfarbe_Nummer"
   Button "Schaltfläche_1" at 863,622 size 149x32; TextOff 'Rollenbahn tippen'
      on Press: SetBit("HochregallagerDB_Motors_Ein")
      on Release: ResetBit("HochregallagerDB_Motors_Ein")
   Rectangle "Rechteck_1" at 886,560 size 96x48
      Appearance <- "HochregallagerDB_Motors_Ein"
   Switch "Schalter_1" at 727,553 size 120x88; CaptionText 'Automatik'; TextOff 'OFF'; TextOn 'ON'
      ProcessValue <- "HochregallagerDB_Automatik"
   Button "Schaltfläche_2" at 751,676 size 236x32; TextOff 'Neue_Palette'
      on Release: ResetBit("HochregallagerDB_Neue_Palette")
      on Press: SetBit("HochregallagerDB_Neue_Palette")
   Rectangle "Rechteck_2" at 102,654 size 69x75
      Visibility <- "Paketempfang_Rollenbahn_DB_Palette_auf_RB1"
   Rectangle "Rechteck_6" at 102,520 size 69x78
      Visibility <- "Paketempfang_Rollenbahn_DB_Palette_auf_RB2"
      Appearance <- "Paketempfang_Rollenbahn_DB_Farbe_RB2"
   Rectangle "Rechteck_7" at 101,378 size 69x88
      Appearance <- "HochregallagerDB_Farbe"
   Rectangle "Rechteck_35" at 162,165 size 47x36
      Appearance <- "HochregallagerDB_Lagerplaetze{19}_Materialfarbe_Nummer"
   Rectangle "Rechteck_8" at 162,216 size 47x36
      Appearance <- "HochregallagerDB_Lagerplaetze{10}_Materialfarbe_Nummer"
   Rectangle "Rechteck_10" at 162,267 size 47x36
      Appearance <- "HochregallagerDB_Lagerplaetze{1}_Materialfarbe_Nummer"
   Rectangle "Rechteck_11" at 224,165 size 47x36
      Appearance <- "HochregallagerDB_Lagerplaetze{20}_Materialfarbe_Nummer"
   Rectangle "Rechteck_12" at 224,216 size 47x36
      Appearance <- "HochregallagerDB_Lagerplaetze{11}_Materialfarbe_Nummer"
   Rectangle "Rechteck_13" at 224,267 size 47x36
      Appearance <- "HochregallagerDB_Lagerplaetze{2}_Materialfarbe_Nummer"
   Rectangle "Rechteck_14" at 286,165 size 47x36
      Appearance <- "HochregallagerDB_Lagerplaetze{21}_Materialfarbe_Nummer"
   Rectangle "Rechteck_15" at 286,216 size 47x36
      Appearance <- "HochregallagerDB_Lagerplaetze{12}_Materialfarbe_Nummer"
   Rectangle "Rechteck_16" at 286,267 size 47x36
      Appearance <- "HochregallagerDB_Lagerplaetze{3}_Materialfarbe_Nummer"
   Rectangle "Rechteck_17" at 348,165 size 47x36
      Appearance <- "HochregallagerDB_Lagerplaetze{22}_Materialfarbe_Nummer"
   Rectangle "Rechteck_18" at 348,216 size 47x36
      Appearance <- "HochregallagerDB_Lagerplaetze{13}_Materialfarbe_Nummer"
   Rectangle "Rechteck_19" at 348,267 size 47x36
      Appearance <- "HochregallagerDB_Lagerplaetze{4}_Materialfarbe_Nummer"
   Rectangle "Rechteck_20" at 410,165 size 47x36
      Appearance <- "HochregallagerDB_Lagerplaetze{23}_Materialfarbe_Nummer"
   Rectangle "Rechteck_21" at 410,216 size 47x36
      Appearance <- "HochregallagerDB_Lagerplaetze{14}_Materialfarbe_Nummer"
   Rectangle "Rechteck_22" at 410,267 size 47x36
      Appearance <- "HochregallagerDB_Lagerplaetze{5}_Materialfarbe_Nummer"
   Rectangle "Rechteck_23" at 472,165 size 47x36
      Appearance <- "HochregallagerDB_Lagerplaetze{24}_Materialfarbe_Nummer"
   Rectangle "Rechteck_24" at 472,216 size 47x36
      Appearance <- "HochregallagerDB_Lagerplaetze{15}_Materialfarbe_Nummer"
   Rectangle "Rechteck_25" at 472,267 size 47x36
      Appearance <- "HochregallagerDB_Lagerplaetze{6}_Materialfarbe_Nummer"
   Rectangle "Rechteck_26" at 534,165 size 47x36
      Appearance <- "HochregallagerDB_Lagerplaetze{25}_Materialfarbe_Nummer"
   Rectangle "Rechteck_27" at 534,216 size 47x36
      Appearance <- "HochregallagerDB_Lagerplaetze{16}_Materialfarbe_Nummer"
   Rectangle "Rechteck_28" at 534,267 size 47x36
      Appearance <- "HochregallagerDB_Lagerplaetze{7}_Materialfarbe_Nummer"
   Rectangle "Rechteck_29" at 596,165 size 47x36
      Appearance <- "HochregallagerDB_Lagerplaetze{26}_Materialfarbe_Nummer"
   Rectangle "Rechteck_30" at 596,216 size 47x36
      Appearance <- "HochregallagerDB_Lagerplaetze{17}_Materialfarbe_Nummer"
   Rectangle "Rechteck_31" at 596,267 size 47x36
      Appearance <- "HochregallagerDB_Lagerplaetze{8}_Materialfarbe_Nummer"
   Rectangle "Rechteck_32" at 658,165 size 47x36
      Appearance <- "HochregallagerDB_Lagerplaetze{27}_Materialfarbe_Nummer"
   Rectangle "Rechteck_33" at 658,216 size 47x36
      Appearance <- "HochregallagerDB_Lagerplaetze{18}_Materialfarbe_Nummer"
   Rectangle "Rechteck_34" at 658,267 size 47x36
      Appearance <- "HochregallagerDB_Lagerplaetze{9}_Materialfarbe_Nummer"
   TextField "Textfeld_2" at 177,276 size 15x22; Text '1'
   TextField "Textfeld_3" at 668,172 size 25x22; Text '27'
   Rectangle "Rechteck_36" at 162,12 size 47x36
      Appearance <- "HochregallagerDB_Lagerplaetze{46}_Materialfarbe_Nummer"
   Rectangle "Rechteck_37" at 162,63 size 47x36
      Appearance <- "HochregallagerDB_Lagerplaetze{37}_Materialfarbe_Nummer"
   Rectangle "Rechteck_38" at 162,114 size 47x36
      Appearance <- "HochregallagerDB_Lagerplaetze{28}_Materialfarbe_Nummer"
   Rectangle "Rechteck_39" at 224,12 size 47x36
      Appearance <- "HochregallagerDB_Lagerplaetze{47}_Materialfarbe_Nummer"
   Rectangle "Rechteck_40" at 224,63 size 47x36
      Appearance <- "HochregallagerDB_Lagerplaetze{38}_Materialfarbe_Nummer"
   Rectangle "Rechteck_41" at 224,114 size 47x36
      Appearance <- "HochregallagerDB_Lagerplaetze{29}_Materialfarbe_Nummer"
   Rectangle "Rechteck_42" at 286,12 size 47x36
      Appearance <- "HochregallagerDB_Lagerplaetze{48}_Materialfarbe_Nummer"
   Rectangle "Rechteck_43" at 286,63 size 47x36
      Appearance <- "HochregallagerDB_Lagerplaetze{39}_Materialfarbe_Nummer"
   Rectangle "Rechteck_44" at 286,114 size 47x36
      Appearance <- "HochregallagerDB_Lagerplaetze{30}_Materialfarbe_Nummer"
   Rectangle "Rechteck_45" at 348,12 size 47x36
      Appearance <- "HochregallagerDB_Lagerplaetze{49}_Materialfarbe_Nummer"
   Rectangle "Rechteck_46" at 348,63 size 47x36
      Appearance <- "HochregallagerDB_Lagerplaetze{40}_Materialfarbe_Nummer"
   Rectangle "Rechteck_47" at 348,114 size 47x36
      Appearance <- "HochregallagerDB_Lagerplaetze{31}_Materialfarbe_Nummer"
   Rectangle "Rechteck_48" at 410,12 size 47x36
      Appearance <- "HochregallagerDB_Lagerplaetze{50}_Materialfarbe_Nummer"
   Rectangle "Rechteck_49" at 410,63 size 47x36
      Appearance <- "HochregallagerDB_Lagerplaetze{41}_Materialfarbe_Nummer"
   Rectangle "Rechteck_50" at 410,114 size 47x36
      Appearance <- "HochregallagerDB_Lagerplaetze{32}_Materialfarbe_Nummer"
   Rectangle "Rechteck_51" at 472,12 size 47x36
      Appearance <- "HochregallagerDB_Lagerplaetze{51}_Materialfarbe_Nummer"
   Rectangle "Rechteck_52" at 472,63 size 47x36
      Appearance <- "HochregallagerDB_Lagerplaetze{42}_Materialfarbe_Nummer"
   Rectangle "Rechteck_53" at 472,114 size 47x36
      Appearance <- "HochregallagerDB_Lagerplaetze{33}_Materialfarbe_Nummer"
   Rectangle "Rechteck_54" at 534,12 size 47x36
      Appearance <- "HochregallagerDB_Lagerplaetze{52}_Materialfarbe_Nummer"
   Rectangle "Rechteck_55" at 534,63 size 47x36
      Appearance <- "HochregallagerDB_Lagerplaetze{43}_Materialfarbe_Nummer"
   Rectangle "Rechteck_56" at 534,114 size 47x36
      Appearance <- "HochregallagerDB_Lagerplaetze{34}_Materialfarbe_Nummer"
   Rectangle "Rechteck_58" at 596,63 size 47x36
      Appearance <- "HochregallagerDB_Lagerplaetze{44}_Materialfarbe_Nummer"
   Rectangle "Rechteck_59" at 596,114 size 47x36
      Appearance <- "HochregallagerDB_Lagerplaetze{35}_Materialfarbe_Nummer"
   Rectangle "Rechteck_60" at 658,12 size 47x36
      Appearance <- "HochregallagerDB_Lagerplaetze{54}_Materialfarbe_Nummer"
   Rectangle "Rechteck_61" at 658,63 size 47x36
      Appearance <- "HochregallagerDB_Lagerplaetze{45}_Materialfarbe_Nummer"
   Rectangle "Rechteck_62" at 658,114 size 47x36
      Appearance <- "HochregallagerDB_Lagerplaetze{36}_Materialfarbe_Nummer"
   TextField "Textfeld_4" at 173,121 size 25x22; Text '28'
   TextField "Textfeld_5" at 668,19 size 25x22; Text '54'
   Rectangle "Rechteck_9" at 114,317 size 34x30
      DirectMovement <- "HochregallagerDB_HMI_X_Bewegung"
      DirectMovement <- "HochregallagerDB_HMI_Z_Bewegung"
      Appearance <- "HochregallagerDB_Stappler_Aktuele_Farbe"
   TextField "Textfeld_1" at 77,320 size 24x22; Text 'ST'
   IOField "EA-Feld_1" at 749,84 size 86x59; FormatPattern 99
      ProcessValue <- "HochregallagerDB_Anzahl_Blau"
   TextField "Textfeld_6" at 746,154 size 98x22; Text 'Anzahl_Blau'
   TextField "Textfeld_7" at 889,154 size 110x22; Text 'Anzahl_Gruen'
   IOField "EA-Feld_2" at 901,84 size 86x59; FormatPattern 99
      ProcessValue <- "HochregallagerDB_Anzahl_Gruen"
   GraphicView "Grafikanzeige_1" at 241,432 size 393x264; Picture "Grafik_1"
   IOField "EA-Feld_4" at 474,631 size 49x30; FormatPattern 99
      ProcessValue <- "HochregallagerDB_Anzahl_Gruen"
   IOField "EA-Feld_3" at 556,632 size 48x29; FormatPattern 99
      ProcessValue <- "HochregallagerDB_Anzahl_Blau"
   Circle "Kreis_1" at 490,492 size 18x18
      Appearance <- "P10_START"
   Circle "Kreis_2" at 532,492 size 18x18
      Appearance <- "P11_STOP"
   Button "Schaltfläche_3" at 480,511 size 38x19; TextOff 'Start'
      on Release: ResetBit("HMI_Eingaben_DB_HMI_Start")
      on Press: SetBit("HMI_Eingaben_DB_HMI_Start")
   Button "Schaltfläche_4" at 522,511 size 38x19; TextOff 'Stop'
      on Release: SetBit("HMI_Eingaben_DB_HMI_Stop")
      on Press: ResetBit("HMI_Eingaben_DB_HMI_Stop")
   Button "Schaltfläche_5" at 308,487 size 37x30; TextOff 'NH'
      on Release: SetBit("HMI_Eingaben_DB_HMI_Not_Halt")
      on Press: ResetBit("HMI_Eingaben_DB_HMI_Not_Halt")
   Switch "Schalter_2" at 307,561 size 50x37; CaptionText 'Switch'; TextOff 'OFF'; TextOn 'ON'
      ProcessValue <- "HMI_Eingaben_DB_HMI_Hauptschalter"
   Rectangle "Rechteck_64" at 570,415 size 23x13
      Appearance <- "P3_MS_GN"
   Rectangle "Rechteck_65" at 570,397 size 23x13
      Appearance <- "P2_MS_GE"
   Rectangle "Rechteck_66" at 570,379 size 23x13
      Appearance <- "P1_MS_RT"
   TextField "Textfeld_9" at 626,382 size 350x44; Text 'Warnschwelle erreicht Nur noch wenige freie Lagerplätze verfügbar.'
      Visibility <- "HochregallagerDB_Warnung_Wenig_Freie_Plaetze"
   TextField "Textfeld_8" at 687,389 size 231x26; Text 'Alle Lagerplaetze sind belegt.'
      Visibility <- "HochregallagerDB_Lager_Voll"
   GraphicView "Grafikanzeige_2" at 366,378 size 63x62; Picture "siren-alert-14183_1024"
      Appearance <- "HochregallagerDB_Stoerung_Aktiv"
   GraphicView "Grafikanzeige_3" at 226,379 size 74x59; Picture "—Pngtree—red warning light long beam_3867061"
      Appearance <- "P12_Anfahrwarnung"
   GraphicView "Grafikanzeige_4" at 28,252 size 74x59; Picture "—Pngtree—red warning light long beam_3867061"
      Appearance <- "P8002_Warnung_Bewegung_2"
   GraphicView "Grafikanzeige_5" at 18,0 size 74x59; Picture "—Pngtree—red warning light long beam_3867061"
      Appearance <- "P8001_Warnung_Bewegung_1"
   IOField "EA-Feld_5" at 820,204 size 86x59; FormatPattern 99
      ProcessValue <- "HochregallagerDB_Anzahl_Unbekannte_Farbe"
   TextField "Textfeld_10" at 786,267 size 147x40; Text 'Anzahl Unbekannte_Farbe'
   TextField "Textfeld_11" at 240,275 size 15x22; Text '2'
   TextField "Textfeld_12" at 177,276 size 15x22; Text '1'
   TextField "Textfeld_13" at 302,274 size 15x22; Text '3'
   TextField "Textfeld_14" at 364,274 size 15x22; Text '4'
   TextField "Textfeld_15" at 426,274 size 15x22; Text '5'
   TextField "Textfeld_16" at 488,273 size 15x22; Text '6'
   TextField "Textfeld_17" at 550,273 size 15x22; Text '7'
   TextField "Textfeld_18" at 610,274 size 15x22; Text '8'
   TextField "Textfeld_19" at 674,273 size 15x22; Text '9'
   TextField "Textfeld_20" at 173,223 size 25x22; Text '10'
   TextField "Textfeld_21" at 234,222 size 25x22; Text '11'
   TextField "Textfeld_22" at 295,222 size 25x22; Text '12'
   TextField "Textfeld_23" at 357,222 size 25x22; Text '13'
   TextField "Textfeld_24" at 420,223 size 25x22; Text '14'
   TextField "Textfeld_25" at 481,222 size 25x22; Text '15'
   TextField "Textfeld_26" at 542,223 size 25x22; Text '16'
   TextField "Textfeld_27" at 604,223 size 25x22; Text '17'
   TextField "Textfeld_28" at 667,223 size 25x22; Text '18'
   TextField "Textfeld_29" at 172,172 size 25x22; Text '19'
   TextField "Textfeld_30" at 234,172 size 25x22; Text '20'
   TextField "Textfeld_31" at 296,172 size 25x22; Text '21'
   TextField "Textfeld_32" at 358,172 size 25x22; Text '22'
   TextField "Textfeld_33" at 420,172 size 25x22; Text '23'
   TextField "Textfeld_34" at 482,172 size 25x22; Text '24'
   TextField "Textfeld_35" at 544,172 size 25x22; Text '25'
   TextField "Textfeld_36" at 606,172 size 25x22; Text '26'
   TextField "Textfeld_37" at 233,121 size 25x22; Text '29'
   TextField "Textfeld_38" at 297,121 size 25x22; Text '30'
   TextField "Textfeld_39" at 359,121 size 25x22; Text '31'
   TextField "Textfeld_40" at 419,121 size 25x22; Text '32'
   TextField "Textfeld_41" at 481,121 size 25x22; Text '33'
   TextField "Textfeld_42" at 545,121 size 25x22; Text '34'
   TextField "Textfeld_43" at 605,121 size 25x22; Text '35'
   TextField "Textfeld_44" at 667,121 size 25x22; Text '36'
   TextField "Textfeld_45" at 171,70 size 25x22; Text '37'
   TextField "Textfeld_46" at 236,70 size 25x22; Text '38'
   TextField "Textfeld_47" at 301,70 size 25x22; Text '39'
   TextField "Textfeld_48" at 360,70 size 25x22; Text '40'
   TextField "Textfeld_49" at 421,70 size 25x22; Text '41'
   TextField "Textfeld_50" at 483,70 size 25x22; Text '42'
   TextField "Textfeld_51" at 545,70 size 25x22; Text '43'
   TextField "Textfeld_52" at 606,70 size 25x22; Text '44'
   TextField "Textfeld_53" at 669,70 size 25x22; Text '45'
   TextField "Textfeld_54" at 173,18 size 25x22; Text '46'
   TextField "Textfeld_55" at 235,18 size 25x22; Text '47'
   TextField "Textfeld_56" at 298,18 size 25x22; Text '48'
   TextField "Textfeld_57" at 361,18 size 25x22; Text '49'
   TextField "Textfeld_58" at 424,18 size 25x22; Text '50'
   TextField "Textfeld_59" at 487,18 size 25x22; Text '51'
   TextField "Textfeld_60" at 550,18 size 25x22; Text '52'
   TextField "Textfeld_61" at 613,18 size 25x22; Text '53'
*)